# EPICS substitutions: db/Beckhoff_2XXX/ecmcEL2262.substitutions
file "ecmcEL2262_binaryOutputArray-chX.template"
{
  pattern {CH_ID}
          {01   }
          {02   }
}

file "ecmcEL2262_common.template"
{
  pattern {}
          {}
}
